Fanuc KAREL source: KT00502.KL

PROGRAM KT00502
%NOLOCKGROUP
VAR
  P1: XYZWPR
  P2: XYZWPR
  OUT: JOINTPOS
BEGIN
  P1.X = 1.0
  P2.Y = 2.0
  P1.X = 1.0
  P2.Y = 2.0
  OUT = P1 : P2
END KT00502
